// TIA Portal V20 export
// export: Created 2026-10-12T15:48:31.6961084Z, ExportSetting WithDefaults, DisplayName Totally Integrated Automation Portal, DisplayVersion V20, DisplayName TIA Portal Openness, DisplayVersion V20, DisplayName TIA Portal Teamcenter Gateway, DisplayVersion V20, DisplayName TIA Portal Version Control Interface, DisplayVersion V20, DisplayName SINAMICS Startdrive Advanced, DisplayVersion V20 SP1 Update 2, DisplayName SINAMICS Startdrive G110M, G120, G120C, G120D, G120P, G115D, DisplayVersion V20 SP1 Update 2, DisplayName SINAMICS Startdrive G130, G150, S120, S150, SINAMICS MV, G220, S200, S210, DisplayVersion V20 SP1 Update 2, DisplayName STEP 7 Professional, DisplayVersion V20, DisplayName STEP 7 Safety, DisplayVersion V20, DisplayName WinCC Basic/Comfort/Advanced, DisplayVersion V20, DisplayName WinCC Professional, DisplayVersion V20, DisplayName WinCC Unified, DisplayVersion V20
FUNCTION "FRK_AlarmHistoryIndex" : Int   // FC40, SCL
{ S7_Optimized_Access := 'TRUE' }
VERSION : 0.1
// Reference-1500 LOCAL_RETAIN: closed history only, keyed by actual Unit scope.
//  No active alarms, commands, sessions or monotonic clocks are restored.
// stored: AutoNumber true, IsIECCheckEnabled false, SetENOAutomatically false, UDAEnableTagReadback false
   VAR_INPUT
      Scope : String;
   END_VAR
BEGIN

   #FRK_AlarmHistoryIndex := 0;
   IF #Scope = 'StationA' THEN
       #FRK_AlarmHistoryIndex := 1;
       RETURN;
   END_IF;
   IF #Scope = 'StationA.Satellite' THEN
       #FRK_AlarmHistoryIndex := 2;
       RETURN;
   END_IF;
   IF #Scope = 'StationB' THEN
       #FRK_AlarmHistoryIndex := 3;
       RETURN;
   END_IF;
END_FUNCTION
